FUNCTION_BLOCK FB_DummyHA IMPLEMENTS I_HigherAuthority, I_LowerAuthority
VAR_INPUT
    ReqAcknowledged : BOOL := TRUE; // Use to control when the HA CHeckRequest Returns TRUE
END_VAR
VAR_OUTPUT
END_VAR
VAR
END_VAR

PROPERTY bLowerAuthorityVetoed : BOOL
GET
END_GET
SET
END_SET
END_PROPERTY

METHOD CheckRequest : BOOL
VAR_INPUT
    nReqID	: DWORD;
END_VAR
CheckRequest := ReqAcknowledged;
END_METHOD

// <Arbiter Internal>
// Elevates the arbitrated BP set to something above.
// Could be another arbiter, or a BP requester/ IO,
// or an FB that locks in a specific portion of the BP set.
METHOD ElevateRequest : BOOL
VAR_INPUT
    HigherAuthority : I_HigherAuthority;
END_VAR
END_METHOD

PROPERTY nLowerAuthorityID : DWORD
GET
nLowerAuthorityID := PMPS_GVL.EXCLUDED_ASSERTION_ID;
END_GET
END_PROPERTY


METHOD RemoveRequest : BOOL
VAR_INPUT
    (*StateID to remove*)
    nReqID	: DWORD;
END_VAR
RemoveRequest := TRUE;
END_METHOD


METHOD RequestBP : BOOL
VAR_INPUT
    (*StateID of state requesting beam parameter set*)
    nReqID	: DWORD;
    (*Requested beam params*)
    stReqBP	: ST_BeamParams;
END_VAR
RequestBP := TRUE;
END_METHOD

END_FUNCTION_BLOCK

(* stored: Version 1.1.0.1
   POU FB_DummyHA: Id {670c3d93-34b2-4592-94f3-5ed3a0dba153}, SpecialFunc None
   Property bLowerAuthorityVetoed: Id {dc69a883-ba74-4f2e-a93f-7cebcc989749}
   Get Get: Id {bf22549d-3b93-41ea-ba39-a97d1feb55bb}
   Set Set: Id {b86c5e73-e5b5-4b68-81a2-72341e89abf1}
   Method CheckRequest: Id {6032c3d9-45c7-4cc0-b102-000af7719efd}
   Method ElevateRequest: Id {f71f404d-56b3-451d-b2b2-c6689b13e32e}
   Property nLowerAuthorityID: Id {32132f8f-263b-4eb5-946b-8283dbd45b0c}
   Get Get: Id {e7806d6e-95f6-4d6c-bc9b-d36d07b4562a}
   Method RemoveRequest: Id {8cc18e1a-c7b1-4978-8d42-4efdc8839d77}
   Method RequestBP: Id {55d2a094-bf30-435f-a214-786bf412cbdf} *)
